(* Logix 5000 project; controller TFF vendor 1 type 14 code 107 rev 33.11; software revision 33.04; part 24 of 38 *)
(* tags used below, declared in another part *)
   Address : DINT;   // Temp Address
   Address2 : DINT;   // Temp Address
   FeedPump_PID_Settings : INT;   // Index
   Index : DINT;   // Index
   result : DINT[2];
   SCL : SCALE;   // Scale Instruction
   TIME : DINT[2];
   AnalogOutput : AnalogOutput[25];   // Analog Output Array
   AnalogPoint : AnalogInput[50];   // Analog Input Array
   ControlLoop : ControlLoop[20];   // Control Loop Array
   ControlLoop_FeedPump : ALIAS FOR ControlLoop[1];
   ControlLoop_PCV101 : ALIAS FOR ControlLoop[3];
   ControlLoop_PCV101_5ms : ALIAS FOR ControlLoop[4];
   ControlLoop_PCV101_RAMP_OUT : REAL;   // Ramp Output
   ControlLoop_PCV201 : ALIAS FOR ControlLoop[5];
   LI101 : ALIAS FOR AnalogPoint[44];
   Mixer : Mixer;   // Mixer config. structure
   PCV101_Control : PCV_Control;   // PCV101 Control UDT
   PumpRunStatus : DINT;   // Pumps Run Status (1 = At least one pump running , 0 = no pump running)
   SIC004 : ALIAS FOR Drive[3];
   SIC004_AO : ALIAS FOR AnalogOutput[5];
   SysControl : SysControl;   // General system status and command
(* Process, continued *)

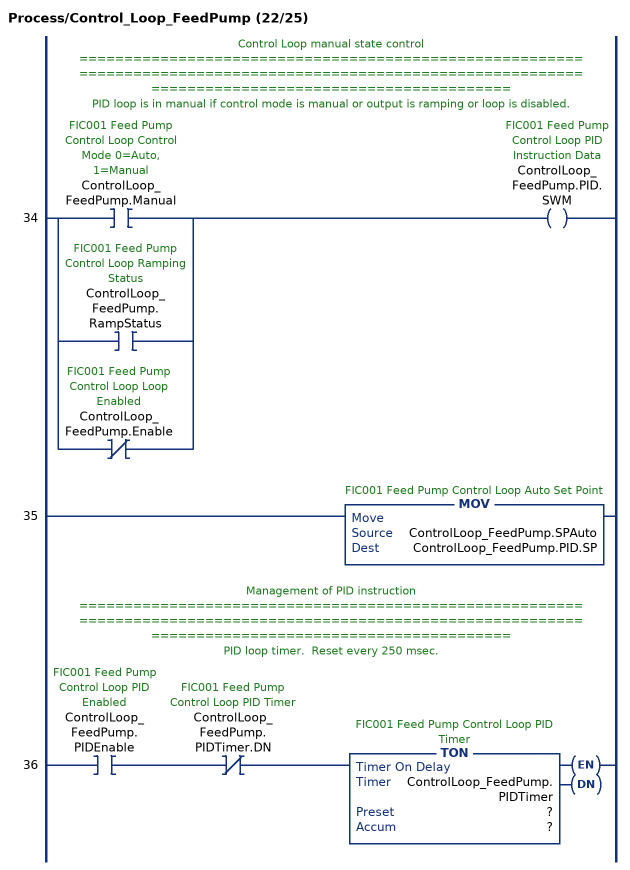
   [picture p191: Process/Control_Loop_FeedPump rungs 34-36]
   // Control Loop manual state control
   // ========================================================================================================================================================
   // PID loop is in manual if control mode is manual or output is ramping or loop is disabled.
   34: [XIC(ControlLoop_FeedPump.Manual) ,XIC(ControlLoop_FeedPump.RampStatus) ,XIO(ControlLoop_FeedPump.Enable) ]OTE(ControlLoop_FeedPump.PID.SWM);
   35: MOV(ControlLoop_FeedPump.SPAuto,ControlLoop_FeedPump.PID.SP);
   // Management of PID instruction
   // ========================================================================================================================================================
   // PID loop timer.  Reset every 250 msec.
   36: XIC(ControlLoop_FeedPump.PIDEnable)XIO(ControlLoop_FeedPump.PIDTimer.DN)TON(ControlLoop_FeedPump.PIDTimer,?,?);
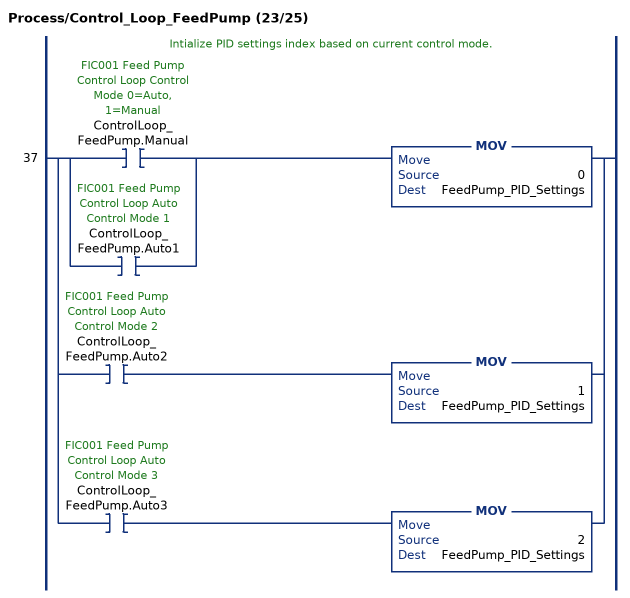
   // Intialize PID settings index based on current control mode.
   37: [[XIC(ControlLoop_FeedPump.Manual) ,XIC(ControlLoop_FeedPump.Auto1) ] MOV(0,FeedPump_PID_Settings) ,XIC(ControlLoop_FeedPump.Auto2) MOV(1,FeedPump_PID_Settings) ,XIC(ControlLoop_FeedPump.Auto3) MOV(2,FeedPump_PID_Settings) ];
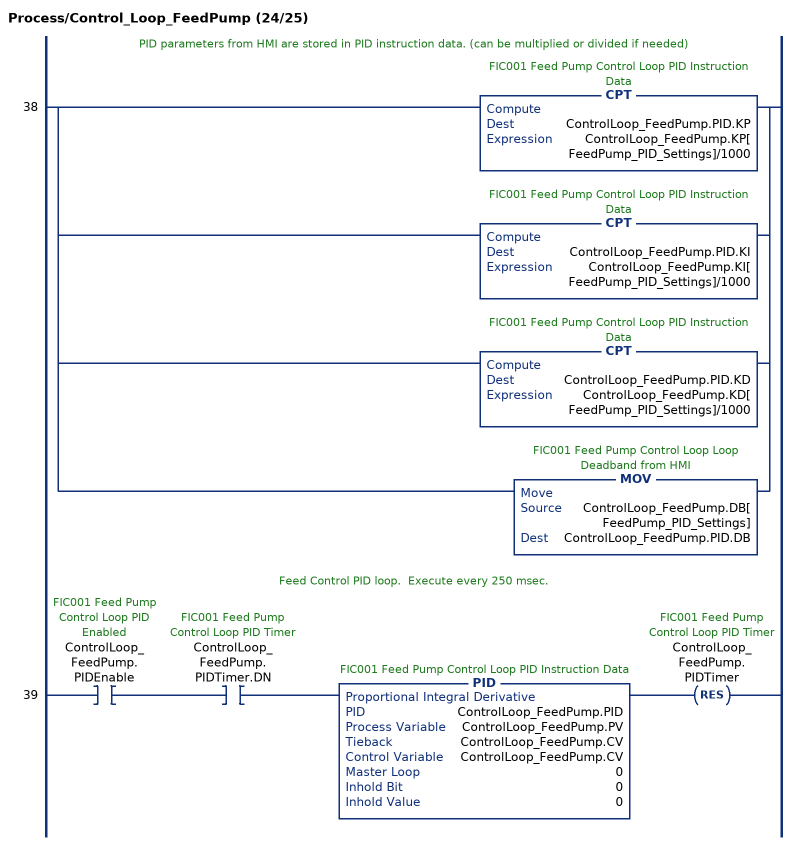
   // PID parameters from HMI are stored in PID instruction data. (can be multiplied or divided if needed)
   38: [CPT(ControlLoop_FeedPump.PID.KP,ControlLoop_FeedPump.KP[FeedPump_PID_Settings]/1000) ,CPT(ControlLoop_FeedPump.PID.KI,ControlLoop_FeedPump.KI[FeedPump_PID_Settings]/1000) ,CPT(ControlLoop_FeedPump.PID.KD,ControlLoop_FeedPump.KD[FeedPump_PID_Settings]/1000) ,MOV(ControlLoop_FeedPump.DB[FeedPump_PID_Settings],ControlLoop_FeedPump.PID.DB) ];
   // Feed Control PID loop.  Execute every 250 msec.
   39: XIC(ControlLoop_FeedPump.PIDEnable)XIC(ControlLoop_FeedPump.PIDTimer.DN)PID(ControlLoop_FeedPump.PID,ControlLoop_FeedPump.PV,ControlLoop_FeedPump.CV,ControlLoop_FeedPump.CV,0,0,0)RES(ControlLoop_FeedPump.PIDTimer);
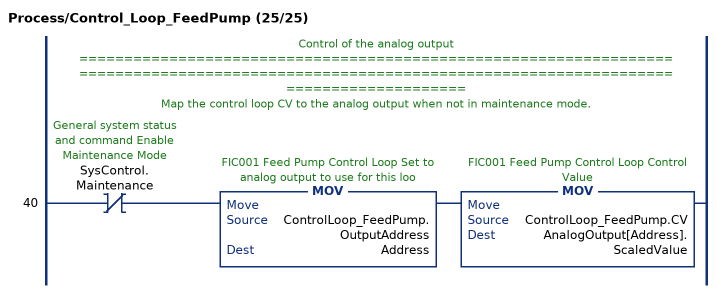
   // Control of the analog output
   // ========================================================================================================================================================
   // Map the control loop CV to the analog output when not in maintenance mode.
   40: XIO(SysControl.Maintenance)MOV(ControlLoop_FeedPump.OutputAddress,Address)MOV(ControlLoop_FeedPump.CV,AnalogOutput[Address].ScaledValue);
END_ROUTINE

ROUTINE Control_Loop_Mixer   (* ladder *)
// Agitator Control Routine
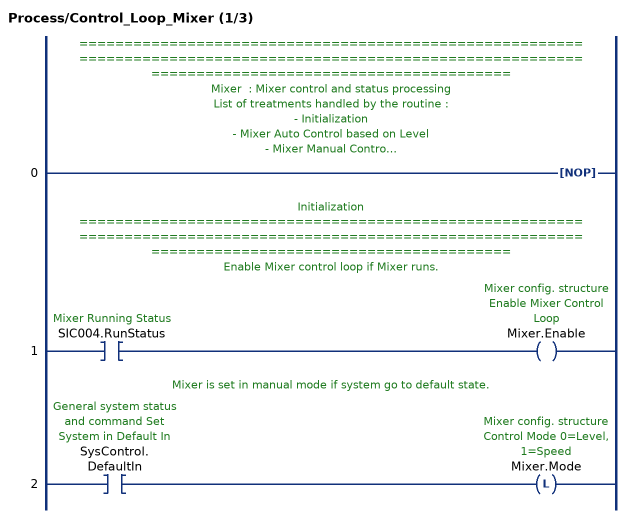
   // ========================================================================================================================================================
   //                                                                                                    Mixer  : Mixer control and status processing
   //                                                     List of treatments handled by the routine :
   //                                                          - Initialization
   //                                                          - Mixer Auto Control based on Level
   //                                                          - Mixer Manual Control
   //                                                     -----------------------------------------------------------------------------------------------------------------------------------------------------
   //                                                     History
   // 		2019-DEC-24 - Merck - Q. Spindler - Initial version for Candidate Release 1.00.00.00.a
   // ========================================================================================================================================================
   0: NOP();
   // Initialization
   // ========================================================================================================================================================
   // Enable Mixer control loop if Mixer runs.
   1: XIC(SIC004.RunStatus)OTE(Mixer.Enable);
   // Mixer is set in manual mode if system go to default state.
   2: XIC(SysControl.DefaultIn)OTL(Mixer.Mode);
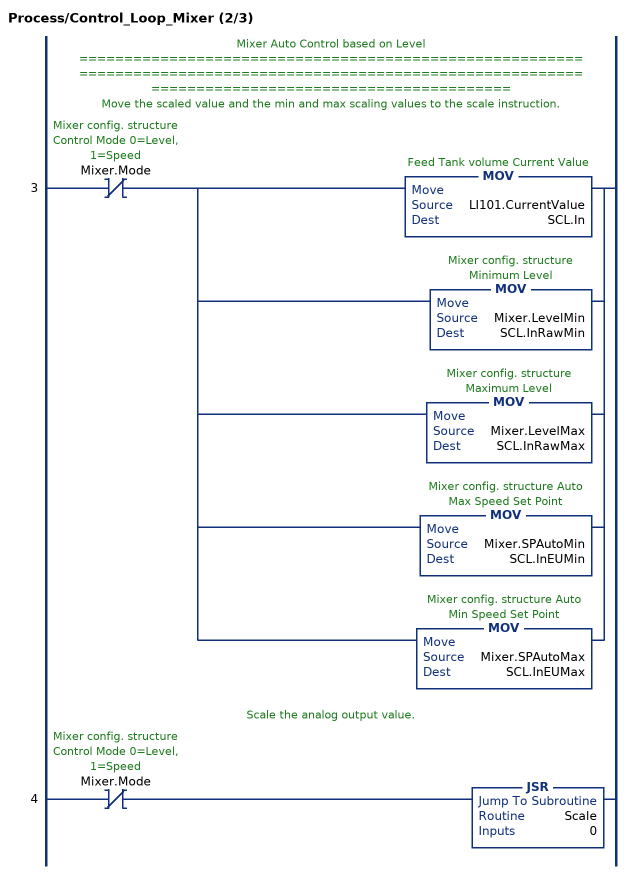
   // Mixer Auto Control based on Level
   // ========================================================================================================================================================
   // Move the scaled value and the min and max scaling values to the scale instruction.
   3: XIO(Mixer.Mode)[MOV(LI101.CurrentValue,SCL.In) ,MOV(Mixer.LevelMin,SCL.InRawMin) ,MOV(Mixer.LevelMax,SCL.InRawMax) ,MOV(Mixer.SPAutoMin,SCL.InEUMin) ,MOV(Mixer.SPAutoMax,SCL.InEUMax) ];
   // Scale the analog output value.
   4: XIO(Mixer.Mode)JSR(Scale,0);
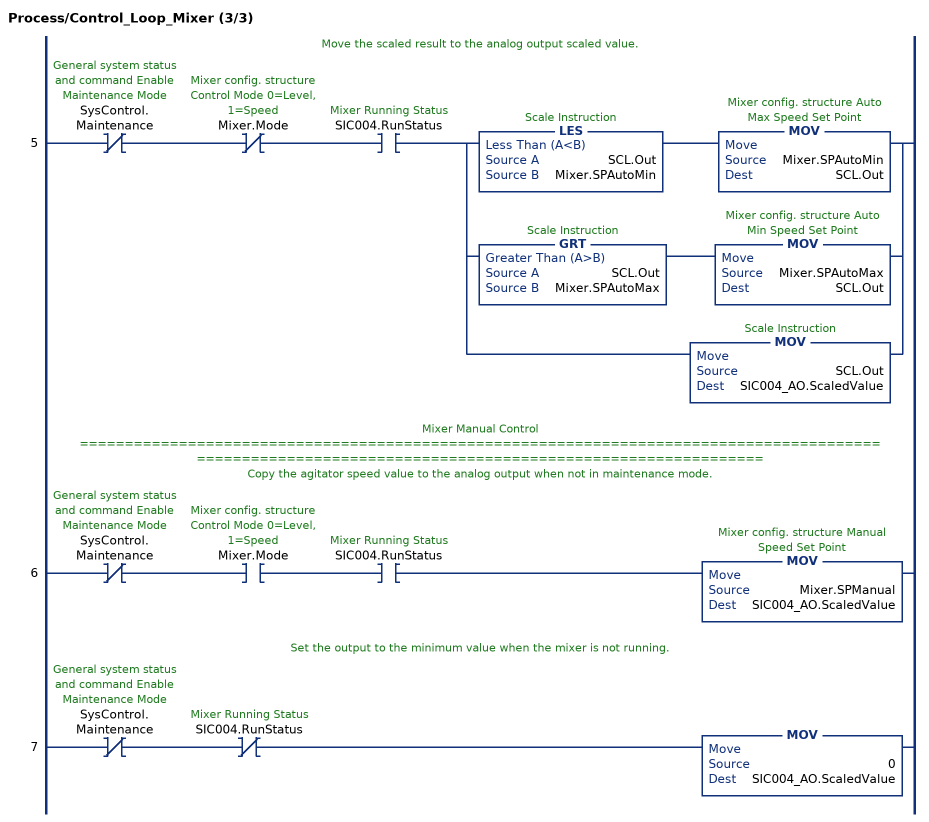
   // Move the scaled result to the analog output scaled value.
   5: XIO(SysControl.Maintenance)XIO(Mixer.Mode)XIC(SIC004.RunStatus)[LES(SCL.Out,Mixer.SPAutoMin) MOV(Mixer.SPAutoMin,SCL.Out) ,GRT(SCL.Out,Mixer.SPAutoMax) MOV(Mixer.SPAutoMax,SCL.Out) ,MOV(SCL.Out,SIC004_AO.ScaledValue) ];
   // Mixer Manual Control
   // ========================================================================================================================================================
   // Copy the agitator speed value to the analog output when not in maintenance mode.
   6: XIO(SysControl.Maintenance)XIC(Mixer.Mode)XIC(SIC004.RunStatus)MOV(Mixer.SPManual,SIC004_AO.ScaledValue);
   // Set the output to the minimum value when the mixer is not running.
   7: XIO(SysControl.Maintenance)XIO(SIC004.RunStatus)MOV(0,SIC004_AO.ScaledValue);
END_ROUTINE

ROUTINE Control_Loop_PCV101   (* ladder *)
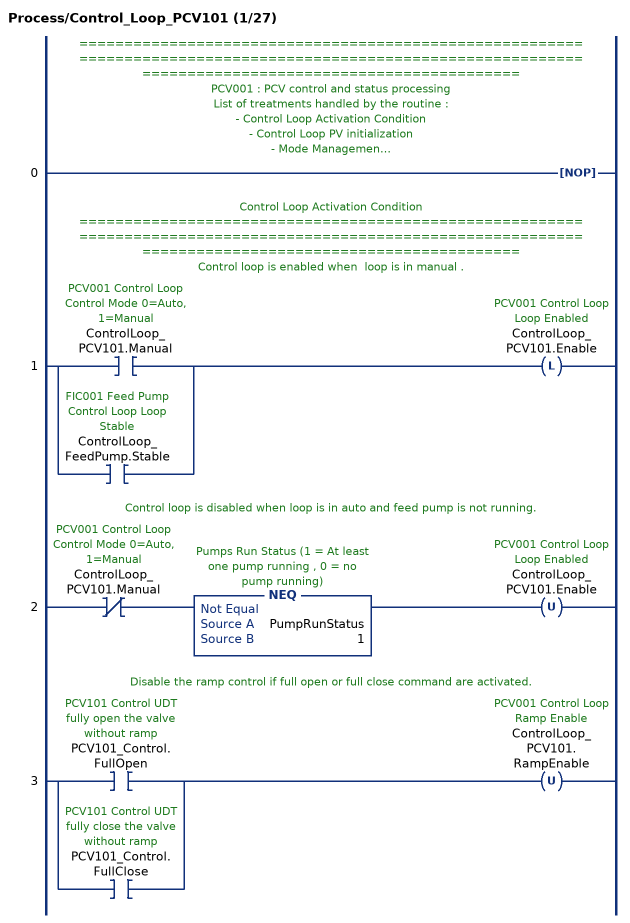
   // ==========================================================================================================================================================
   //                                                  PCV001 : PCV control and status processing
   //                                                     List of treatments handled by the routine :
   //                                                          - Control Loop Activation Condition
   //                                                  - Control Loop PV initialization
   //                                                - Mode Management
   //                                                        - Control Loop Setpoint management
   //                                                        - Control Loop deadband calculation
   //                                                          - Management of ramping control
   //                                                          - Control Loop Stability control
   //                                                          - Full Open - Full Close processing
   //                                                          - Management of PID instruction
   //                                                          - Control of the analog output
   //                                                     -----------------------------------------------------------------------------------------------------------------------------------------------------
   //                                                     History
   // 		2019-DEC-24 - Merck - Q. Spindler - Initial version for Candidate Release 1.00.00.00.a
   // 		2020-SEP-09 - Merck - Q. Spindler - Modifications for Candidate Release 1.00.00.00.d
   // 					- Add ControlLoop Enable and not manual condition for DBOK status
   // 		2021-APR-16 - Merck - Q. Spindler - Modifications for Candidate Release 1.00.00.00.e
   //                                        - Add Initialize address if no mode selected.
   // ==========================================================================================================================================================
   0: NOP();
   // Control Loop Activation Condition
   // ==========================================================================================================================================================
   // Control loop is enabled when  loop is in manual .
   1: [XIC(ControlLoop_PCV101.Manual) ,XIC(ControlLoop_FeedPump.Stable) ]OTL(ControlLoop_PCV101.Enable);
   // Control loop is disabled when loop is in auto and feed pump is not running.
   2: XIO(ControlLoop_PCV101.Manual)NEQ(PumpRunStatus,1)OTU(ControlLoop_PCV101.Enable);
   // Disable the ramp control if full open or full close command are activated.
   3: [XIC(PCV101_Control.FullOpen) ,XIC(PCV101_Control.FullClose) ]OTU(ControlLoop_PCV101.RampEnable);
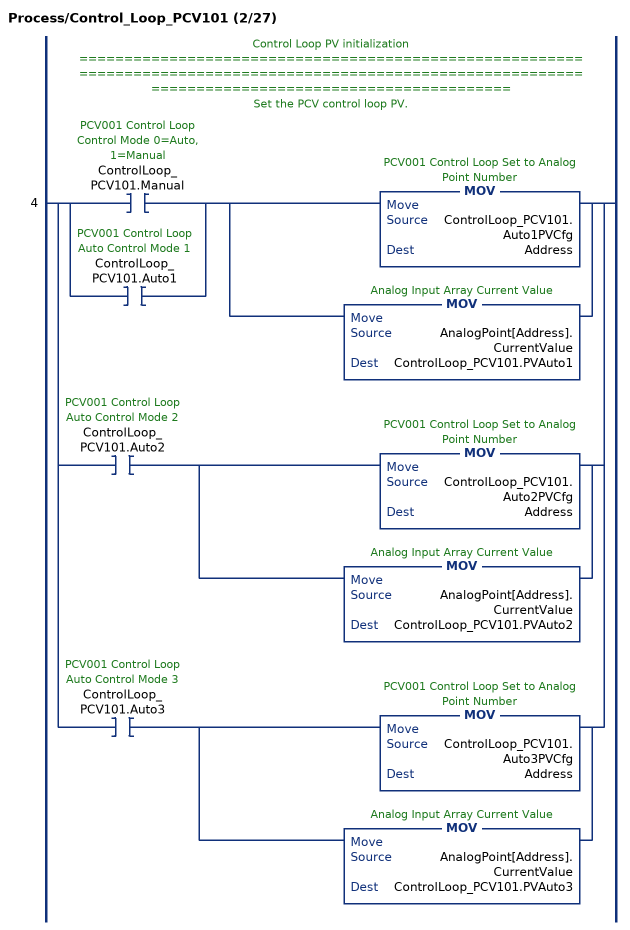
   // Control Loop PV initialization
   // ========================================================================================================================================================
   // Set the PCV control loop PV.
   4: [[[XIC(ControlLoop_PCV101.Manual) ,XIC(ControlLoop_PCV101.Auto1) ] [MOV(ControlLoop_PCV101.Auto1PVCfg,Address) ,MOV(AnalogPoint[Address].CurrentValue,ControlLoop_PCV101.PVAuto1) ] ,XIC(ControlLoop_PCV101.Auto2) [MOV(ControlLoop_PCV101.Auto2PVCfg,Address) ,MOV(AnalogPoint[Address].CurrentValue,ControlLoop_PCV101.PVAuto2) ] ] ,XIC(ControlLoop_PCV101.Auto3) [MOV(ControlLoop_PCV101.Auto3PVCfg,Address) ,MOV(AnalogPoint[Address].CurrentValue,ControlLoop_PCV101.PVAuto3) ] ];
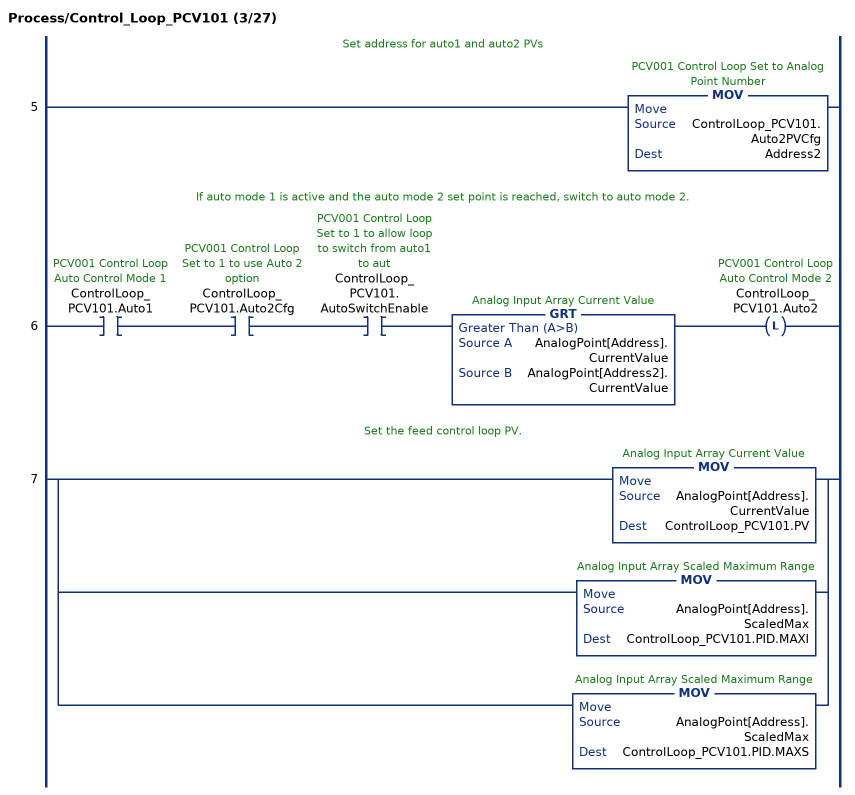
   // Set address for auto1 and auto2 PVs
   5: MOV(ControlLoop_PCV101.Auto2PVCfg,Address2);
   // If auto mode 1 is active and the auto mode 2 set point is reached, switch to auto mode 2.
   6: XIC(ControlLoop_PCV101.Auto1)XIC(ControlLoop_PCV101.Auto2Cfg)XIC(ControlLoop_PCV101.AutoSwitchEnable)GRT(AnalogPoint[Address].CurrentValue,AnalogPoint[Address2].CurrentValue)OTL(ControlLoop_PCV101.Auto2);
   // Set the feed control loop PV.
   7: [MOV(AnalogPoint[Address].CurrentValue,ControlLoop_PCV101.PV) ,MOV(AnalogPoint[Address].ScaledMax,ControlLoop_PCV101.PID.MAXI) ,MOV(AnalogPoint[Address].ScaledMax,ControlLoop_PCV101.PID.MAXS) ];
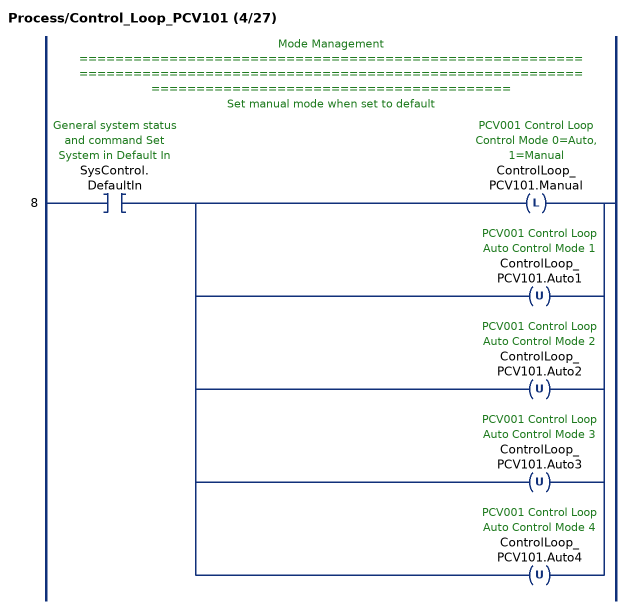
   // Mode Management
   // ========================================================================================================================================================
   // Set manual mode when set to default
   8: XIC(SysControl.DefaultIn)[OTL(ControlLoop_PCV101.Manual) ,OTU(ControlLoop_PCV101.Auto1) ,OTU(ControlLoop_PCV101.Auto2) ,OTU(ControlLoop_PCV101.Auto3) ,OTU(ControlLoop_PCV101.Auto4) ];
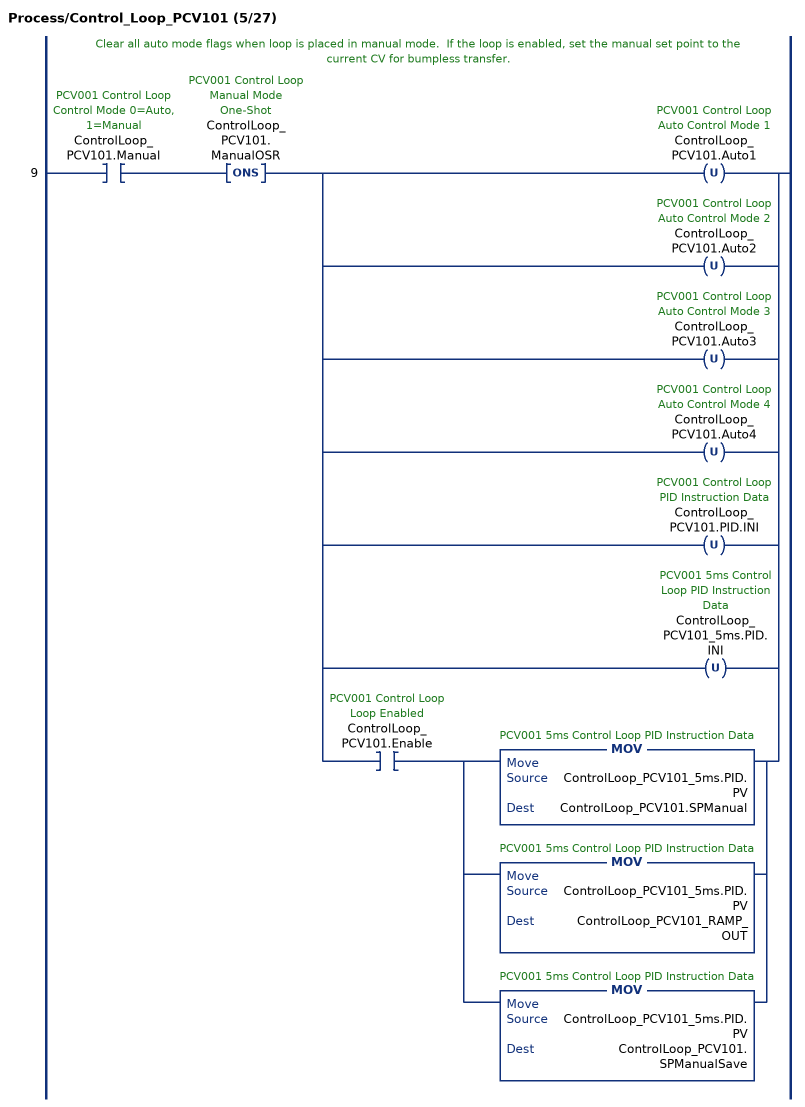
   // Clear all auto mode flags when loop is placed in manual mode.  If the loop is enabled, set the manual set point to the current CV for bumpless transfer.
   9: XIC(ControlLoop_PCV101.Manual)ONS(ControlLoop_PCV101.ManualOSR)[OTU(ControlLoop_PCV101.Auto1) ,OTU(ControlLoop_PCV101.Auto2) ,OTU(ControlLoop_PCV101.Auto3) ,OTU(ControlLoop_PCV101.Auto4) ,OTU(ControlLoop_PCV101.PID.INI) ,OTU(ControlLoop_PCV101_5ms.PID.INI) ,XIC(ControlLoop_PCV101.Enable) [MOV(ControlLoop_PCV101_5ms.PID.PV,ControlLoop_PCV101.SPManual) ,MOV(ControlLoop_PCV101_5ms.PID.PV,ControlLoop_PCV101_RAMP_OUT) ,MOV(ControlLoop_PCV101_5ms.PID.PV,ControlLoop_PCV101.SPManualSave) ] ];
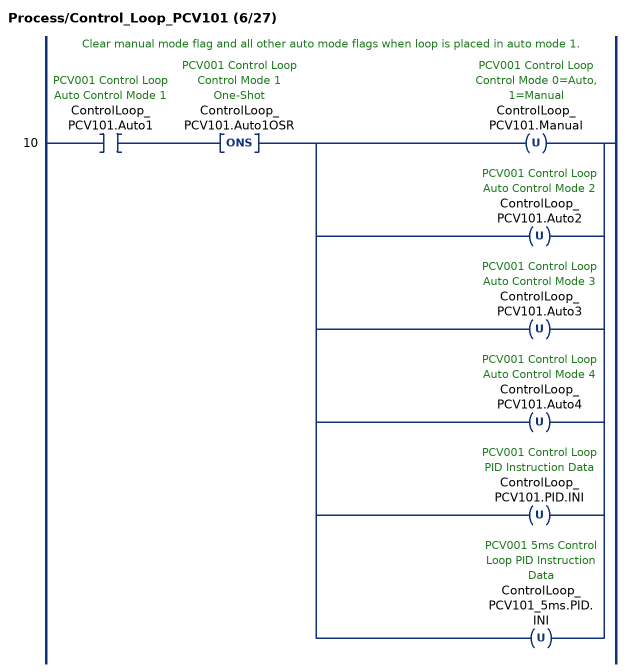
   // Clear manual mode flag and all other auto mode flags when loop is placed in auto mode 1.
   10: XIC(ControlLoop_PCV101.Auto1)ONS(ControlLoop_PCV101.Auto1OSR)[OTU(ControlLoop_PCV101.Manual) ,OTU(ControlLoop_PCV101.Auto2) ,OTU(ControlLoop_PCV101.Auto3) ,OTU(ControlLoop_PCV101.Auto4) ,OTU(ControlLoop_PCV101.PID.INI) ,OTU(ControlLoop_PCV101_5ms.PID.INI) ];
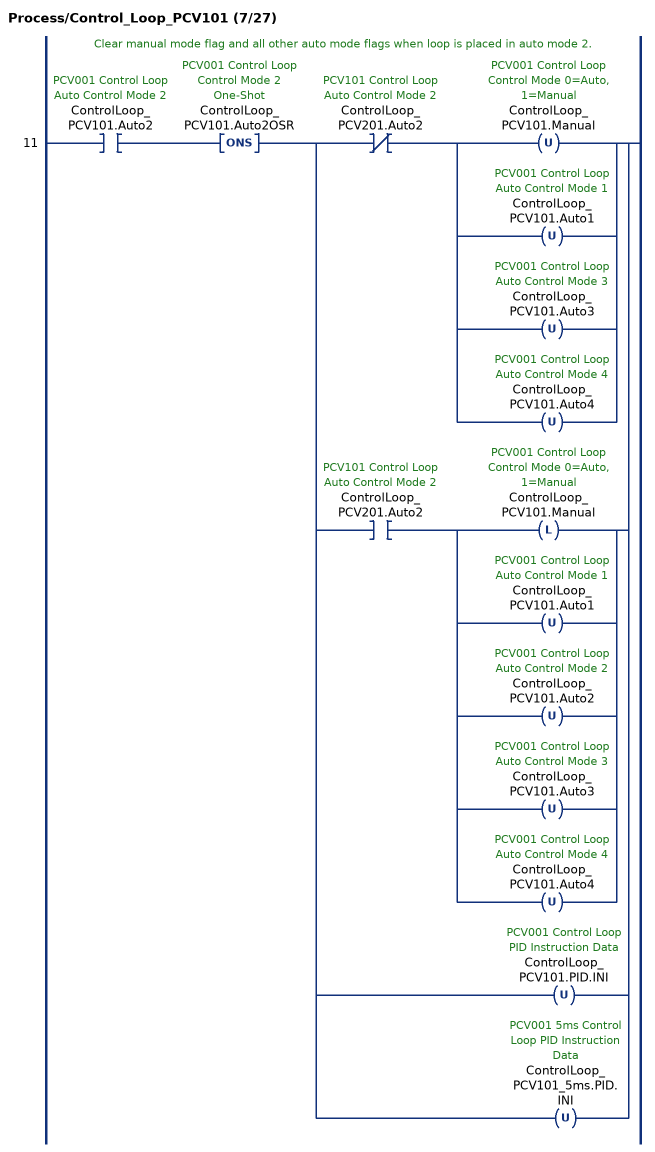
   // Clear manual mode flag and all other auto mode flags when loop is placed in auto mode 2.
   11: XIC(ControlLoop_PCV101.Auto2)ONS(ControlLoop_PCV101.Auto2OSR)[XIO(ControlLoop_PCV201.Auto2) [OTU(ControlLoop_PCV101.Manual) ,OTU(ControlLoop_PCV101.Auto1) ,OTU(ControlLoop_PCV101.Auto3) ,OTU(ControlLoop_PCV101.Auto4) ] ,XIC(ControlLoop_PCV201.Auto2) [OTL(ControlLoop_PCV101.Manual) ,OTU(ControlLoop_PCV101.Auto1) ,OTU(ControlLoop_PCV101.Auto2) ,OTU(ControlLoop_PCV101.Auto3) ,OTU(ControlLoop_PCV101.Auto4) ] ,OTU(ControlLoop_PCV101.PID.INI) ,OTU(ControlLoop_PCV101_5ms.PID.INI) ];
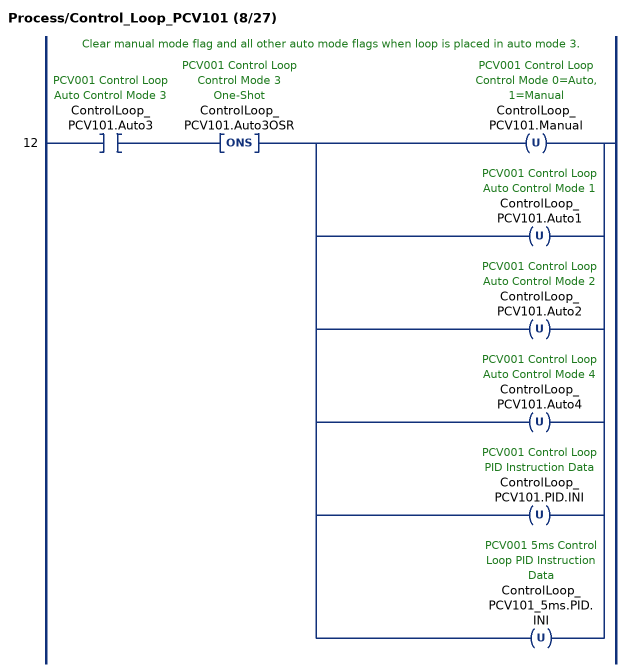
   // Clear manual mode flag and all other auto mode flags when loop is placed in auto mode 3.
   12: XIC(ControlLoop_PCV101.Auto3)ONS(ControlLoop_PCV101.Auto3OSR)[OTU(ControlLoop_PCV101.Manual) ,OTU(ControlLoop_PCV101.Auto1) ,OTU(ControlLoop_PCV101.Auto2) ,OTU(ControlLoop_PCV101.Auto4) ,OTU(ControlLoop_PCV101.PID.INI) ,OTU(ControlLoop_PCV101_5ms.PID.INI) ];
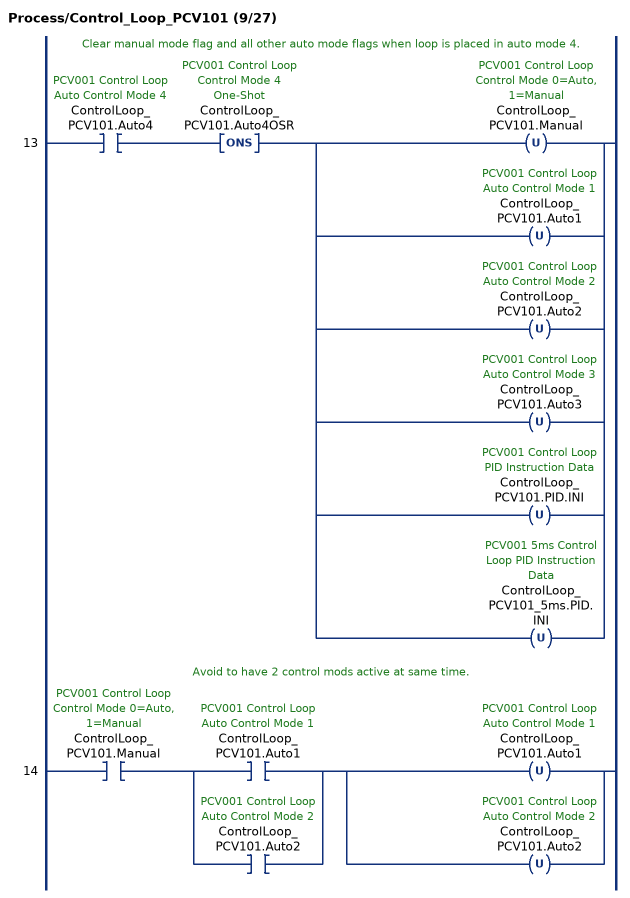
   // Clear manual mode flag and all other auto mode flags when loop is placed in auto mode 4.
   13: XIC(ControlLoop_PCV101.Auto4)ONS(ControlLoop_PCV101.Auto4OSR)[OTU(ControlLoop_PCV101.Manual) ,OTU(ControlLoop_PCV101.Auto1) ,OTU(ControlLoop_PCV101.Auto2) ,OTU(ControlLoop_PCV101.Auto3) ,OTU(ControlLoop_PCV101.PID.INI) ,OTU(ControlLoop_PCV101_5ms.PID.INI) ];
   // Avoid to have 2 control mods active at same time.
   14: XIC(ControlLoop_PCV101.Manual)[XIC(ControlLoop_PCV101.Auto1) ,XIC(ControlLoop_PCV101.Auto2) ][OTU(ControlLoop_PCV101.Auto1) ,OTU(ControlLoop_PCV101.Auto2) ];
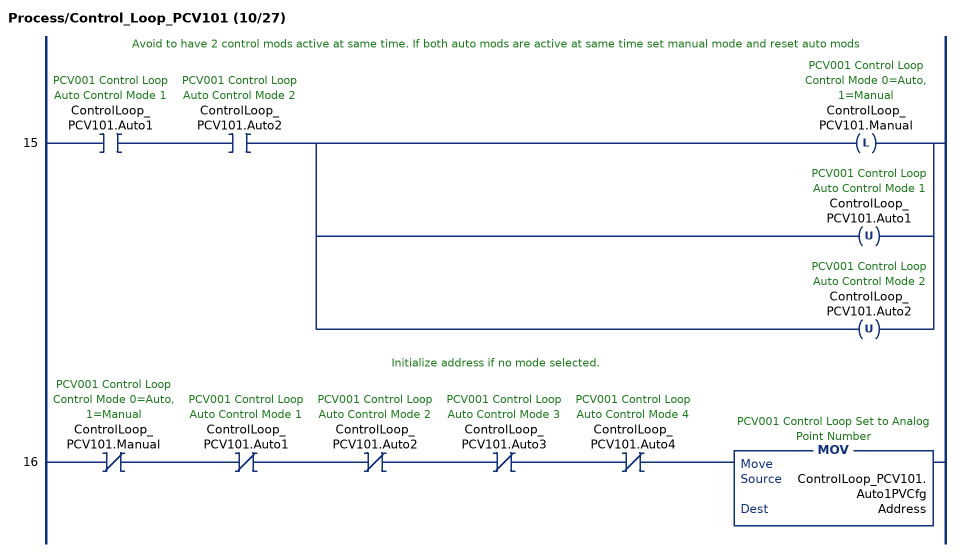
   // Avoid to have 2 control mods active at same time. If both auto mods are active at same time set manual mode and reset auto mods
   15: XIC(ControlLoop_PCV101.Auto1)XIC(ControlLoop_PCV101.Auto2)[OTL(ControlLoop_PCV101.Manual) ,OTU(ControlLoop_PCV101.Auto1) ,OTU(ControlLoop_PCV101.Auto2) ];
   // Initialize address if no mode selected.
   16: XIO(ControlLoop_PCV101.Manual)XIO(ControlLoop_PCV101.Auto1)XIO(ControlLoop_PCV101.Auto2)XIO(ControlLoop_PCV101.Auto3)XIO(ControlLoop_PCV101.Auto4)MOV(ControlLoop_PCV101.Auto1PVCfg,Address);
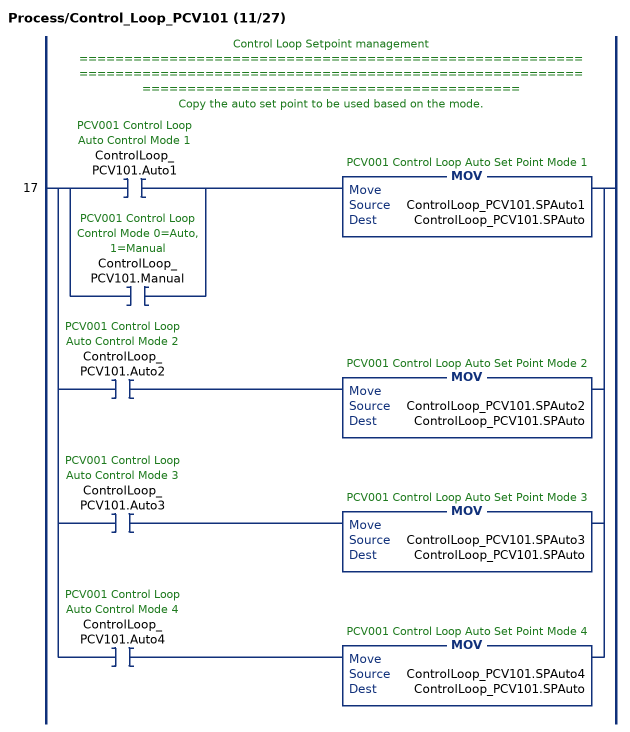
   // Control Loop Setpoint management
   // ==========================================================================================================================================================
   // Copy the auto set point to be used based on the mode.
   17: [[XIC(ControlLoop_PCV101.Auto1) ,XIC(ControlLoop_PCV101.Manual) ] MOV(ControlLoop_PCV101.SPAuto1,ControlLoop_PCV101.SPAuto) ,XIC(ControlLoop_PCV101.Auto2) MOV(ControlLoop_PCV101.SPAuto2,ControlLoop_PCV101.SPAuto) ,XIC(ControlLoop_PCV101.Auto3) MOV(ControlLoop_PCV101.SPAuto3,ControlLoop_PCV101.SPAuto) ,XIC(ControlLoop_PCV101.Auto4) MOV(ControlLoop_PCV101.SPAuto4,ControlLoop_PCV101.SPAuto) ];
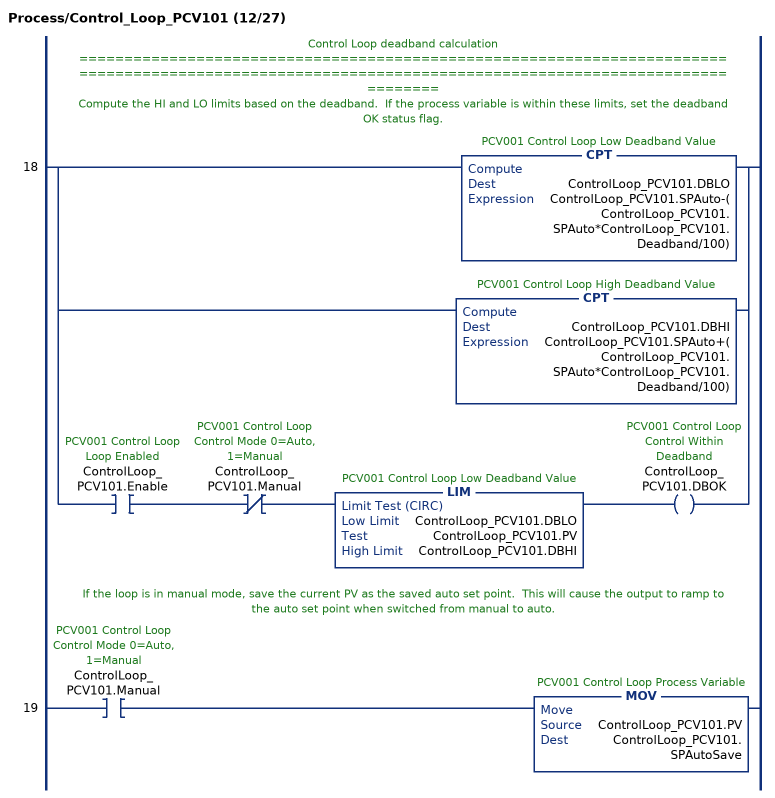
   // Control Loop deadband calculation
   // ========================================================================================================================================================
   // Compute the HI and LO limits based on the deadband.  If the process variable is within these limits, set the deadband OK status flag.
   18: [CPT(ControlLoop_PCV101.DBLO,ControlLoop_PCV101.SPAuto-(ControlLoop_PCV101.SPAuto*ControlLoop_PCV101.Deadband/100)) ,CPT(ControlLoop_PCV101.DBHI,ControlLoop_PCV101.SPAuto+(ControlLoop_PCV101.SPAuto*ControlLoop_PCV101.Deadband/100)) ,XIC(ControlLoop_PCV101.Enable) XIO(ControlLoop_PCV101.Manual) LIM(ControlLoop_PCV101.DBLO,ControlLoop_PCV101.PV,ControlLoop_PCV101.DBHI) OTE(ControlLoop_PCV101.DBOK) ];
   // If the loop is in manual mode, save the current PV as the saved auto set point.  This will cause the output to ramp to the auto set point when switched from manual to auto.
   19: XIC(ControlLoop_PCV101.Manual)MOV(ControlLoop_PCV101.PV,ControlLoop_PCV101.SPAutoSave);
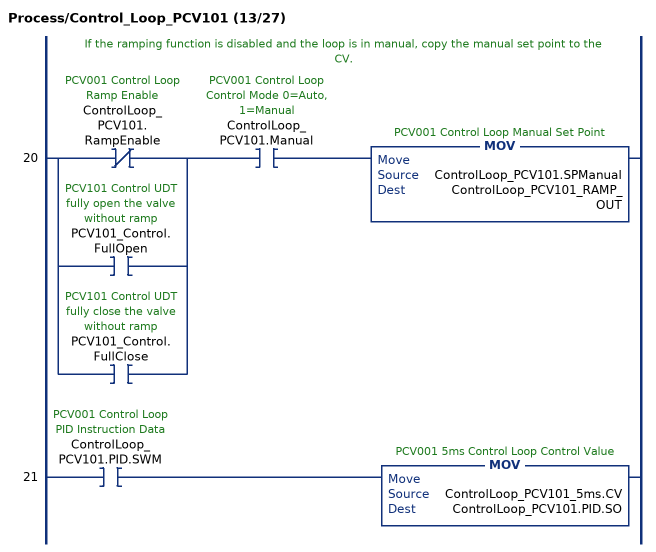
   // If the ramping function is disabled and the loop is in manual, copy the manual set point to the CV.
   20: [XIO(ControlLoop_PCV101.RampEnable) ,XIC(PCV101_Control.FullOpen) ,XIC(PCV101_Control.FullClose) ]XIC(ControlLoop_PCV101.Manual)MOV(ControlLoop_PCV101.SPManual,ControlLoop_PCV101_RAMP_OUT);
   21: XIC(ControlLoop_PCV101.PID.SWM)MOV(ControlLoop_PCV101_5ms.CV,ControlLoop_PCV101.PID.SO);
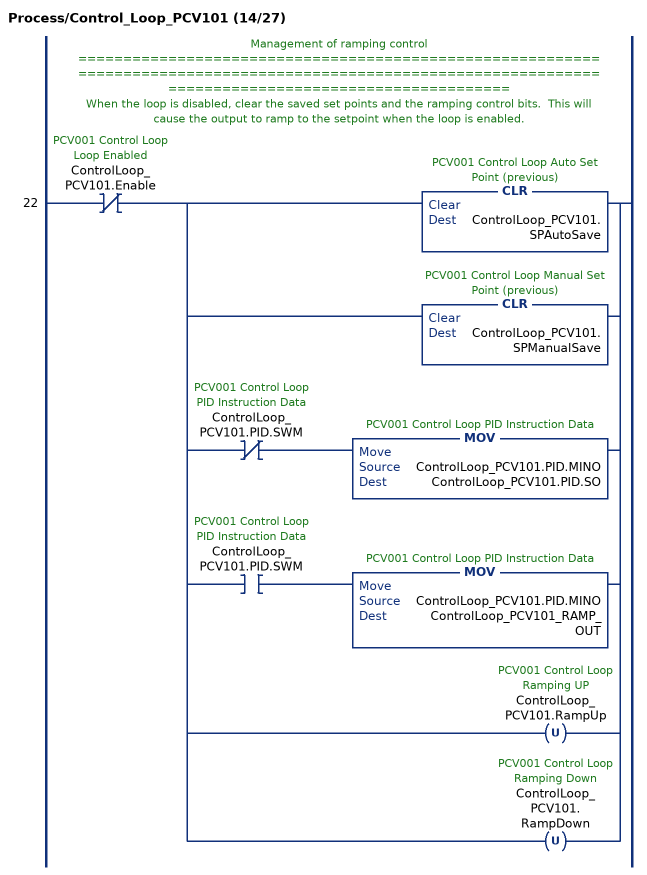
   // Management of ramping control
   // ==========================================================================================================================================================
   // When the loop is disabled, clear the saved set points and the ramping control bits.  This will cause the output to ramp to the setpoint when the loop is enabled.
   22: XIO(ControlLoop_PCV101.Enable)[CLR(ControlLoop_PCV101.SPAutoSave) ,CLR(ControlLoop_PCV101.SPManualSave) ,XIO(ControlLoop_PCV101.PID.SWM) MOV(ControlLoop_PCV101.PID.MINO,ControlLoop_PCV101.PID.SO) ,XIC(ControlLoop_PCV101.PID.SWM) MOV(ControlLoop_PCV101.PID.MINO,ControlLoop_PCV101_RAMP_OUT) ,OTU(ControlLoop_PCV101.RampUp) ,OTU(ControlLoop_PCV101.RampDown) ];
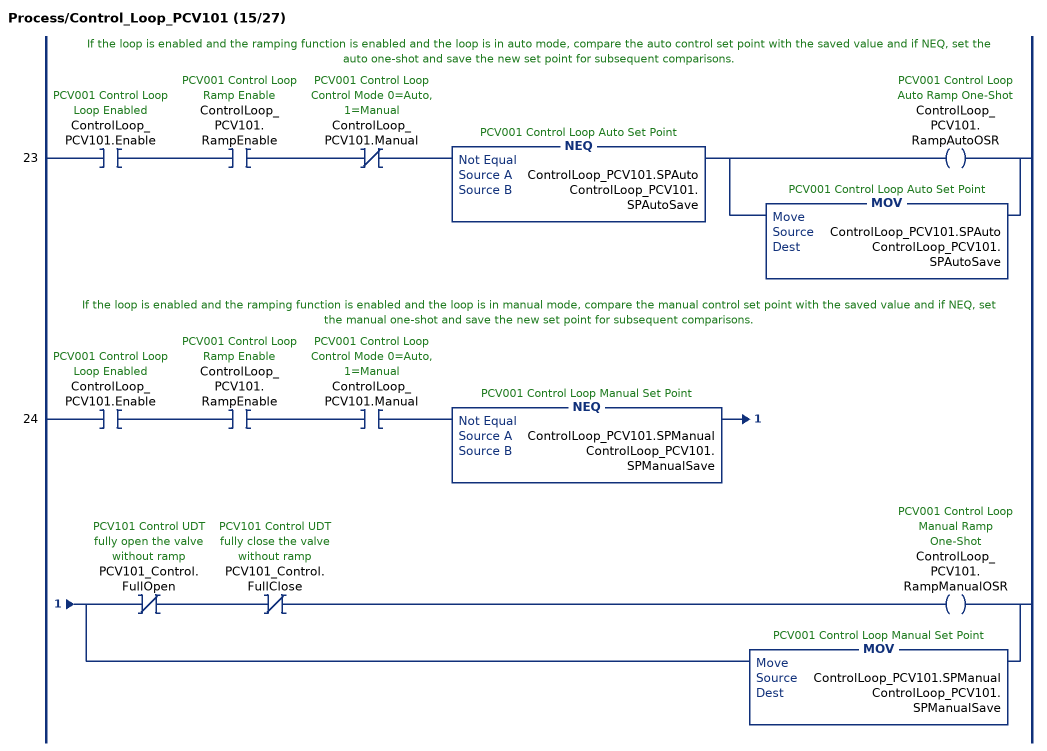
   // If the loop is enabled and the ramping function is enabled and the loop is in auto mode, compare the auto control set point with the saved value and if NEQ, set the auto one-shot and save the new set point for subsequent comparisons.
   23: XIC(ControlLoop_PCV101.Enable)XIC(ControlLoop_PCV101.RampEnable)XIO(ControlLoop_PCV101.Manual)NEQ(ControlLoop_PCV101.SPAuto,ControlLoop_PCV101.SPAutoSave)[OTE(ControlLoop_PCV101.RampAutoOSR) ,MOV(ControlLoop_PCV101.SPAuto,ControlLoop_PCV101.SPAutoSave) ];
   // If the loop is enabled and the ramping function is enabled and the loop is in manual mode, compare the manual control set point with the saved value and if NEQ, set the manual one-shot and save the new set point for subsequent comparisons.
   24: XIC(ControlLoop_PCV101.Enable)XIC(ControlLoop_PCV101.RampEnable)XIC(ControlLoop_PCV101.Manual)NEQ(ControlLoop_PCV101.SPManual,ControlLoop_PCV101.SPManualSave)[XIO(PCV101_Control.FullOpen) XIO(PCV101_Control.FullClose) OTE(ControlLoop_PCV101.RampManualOSR) ,MOV(ControlLoop_PCV101.SPManual,ControlLoop_PCV101.SPManualSave) ];
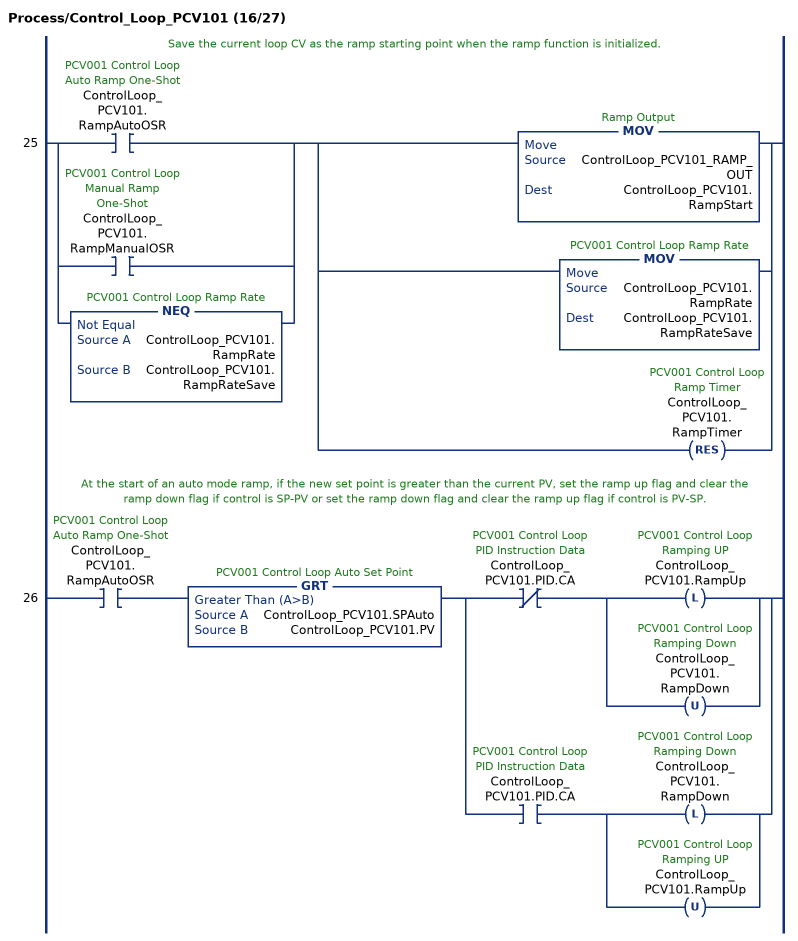
   // Save the current loop CV as the ramp starting point when the ramp function is initialized.
   25: [XIC(ControlLoop_PCV101.RampAutoOSR) ,XIC(ControlLoop_PCV101.RampManualOSR) ,NEQ(ControlLoop_PCV101.RampRate,ControlLoop_PCV101.RampRateSave) ][MOV(ControlLoop_PCV101_RAMP_OUT,ControlLoop_PCV101.RampStart) ,MOV(ControlLoop_PCV101.RampRate,ControlLoop_PCV101.RampRateSave) ,RES(ControlLoop_PCV101.RampTimer) ];
   // At the start of an auto mode ramp, if the new set point is greater than the current PV, set the ramp up flag and clear the ramp down flag if control is SP-PV or set the ramp down flag and clear the ramp up flag if control is PV-SP.
   26: XIC(ControlLoop_PCV101.RampAutoOSR)GRT(ControlLoop_PCV101.SPAuto,ControlLoop_PCV101.PV)[XIO(ControlLoop_PCV101.PID.CA) [OTL(ControlLoop_PCV101.RampUp) ,OTU(ControlLoop_PCV101.RampDown) ] ,XIC(ControlLoop_PCV101.PID.CA) [OTL(ControlLoop_PCV101.RampDown) ,OTU(ControlLoop_PCV101.RampUp) ] ];
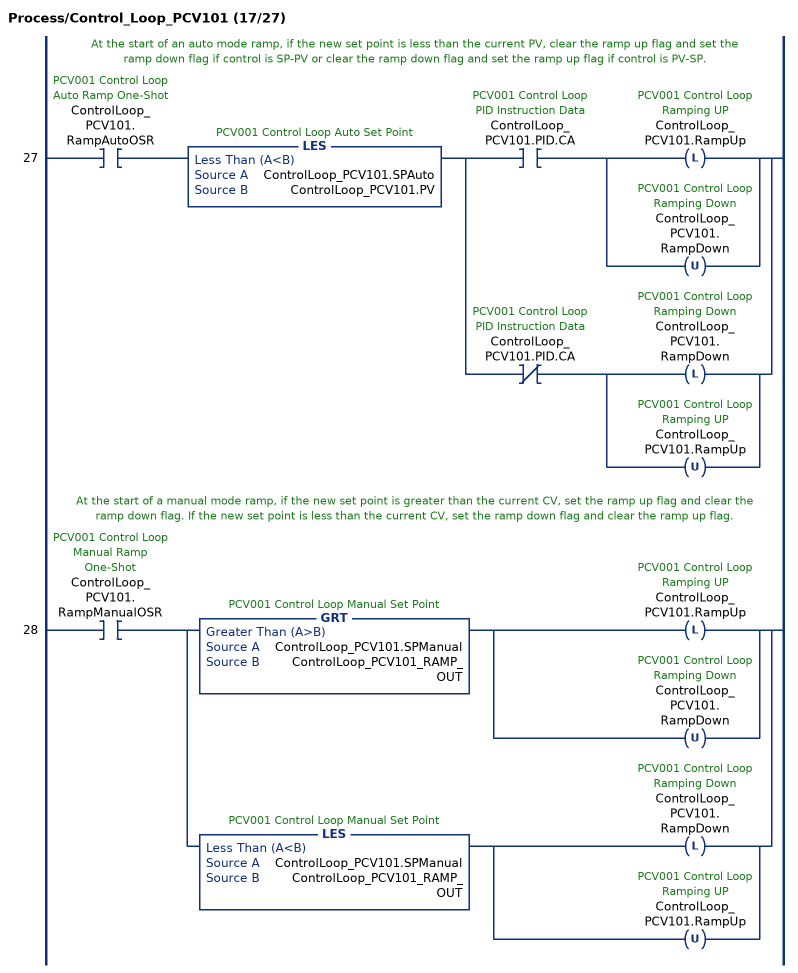
   // At the start of an auto mode ramp, if the new set point is less than the current PV, clear the ramp up flag and set the ramp down flag if control is SP-PV or clear the ramp down flag and set the ramp up flag if control is PV-SP.
   27: XIC(ControlLoop_PCV101.RampAutoOSR)LES(ControlLoop_PCV101.SPAuto,ControlLoop_PCV101.PV)[XIC(ControlLoop_PCV101.PID.CA) [OTL(ControlLoop_PCV101.RampUp) ,OTU(ControlLoop_PCV101.RampDown) ] ,XIO(ControlLoop_PCV101.PID.CA) [OTL(ControlLoop_PCV101.RampDown) ,OTU(ControlLoop_PCV101.RampUp) ] ];
   // At the start of a manual mode ramp, if the new set point is greater than the current CV, set the ramp up flag and clear the ramp down flag. If the new set point is less than the current CV, set the ramp down flag and clear the ramp up flag.
   28: XIC(ControlLoop_PCV101.RampManualOSR)[GRT(ControlLoop_PCV101.SPManual,ControlLoop_PCV101_RAMP_OUT) [OTL(ControlLoop_PCV101.RampUp) ,OTU(ControlLoop_PCV101.RampDown) ] ,LES(ControlLoop_PCV101.SPManual,ControlLoop_PCV101_RAMP_OUT) [OTL(ControlLoop_PCV101.RampDown) ,OTU(ControlLoop_PCV101.RampUp) ] ];
